(* IEC 61131-3 sources: JingjiangArm/moonboxpro_arm_8.4/Application/Application/任务列表/ExtTask/动作处理/油墨槽控制, 9 files *)

(* ---- StInkGrooveCtl.st ---- *)
(*@CES
Name=StInkGrooveCtl
Type=Gvl
TypeGuid=2db5746d-d284-4425-9f7f-2663a34b0ebc
Guid=c6ce6a04-2efb-4550-ab95-73592a3e1ea7
HasDeclaration=True
HasImplementation=False
*)
{DECLARATION}
TYPE StInkGrooveCtl :(*油墨槽控制@不保持|50bytes*)
STRUCT
	bySts							:BYTE;(*状态@就不用枚举了*)
	byMovingSts						:BYTE;(*运动状态|=0 不运动|=1 上升|=2 下降*)
	xCtlMode						:BOOL;(*控制模式|=false速度模式|=true 位置模式*)
	xMoveDir						:BOOL;(*运动的方向*)
	rVel							:REAL;(*速度值@r/min*)
	rMoveDis						:REAL;(*需要运动的距离@mm(带方向)*)
	diMoveDis_Pulse					:DINT;(*需要运动的距离(正值)@pulse*)
	wLastPulse_Act_Rd				:WORD;(*实际读取的脉冲数记录@上一拍*)
	xZeroValid						:BOOL;(*零位有效*)
	diPulse_Moved					:DINT;(*已经移动的脉冲|在原点处会更新为0*)
	rPos_Cur						:REAL;(*当前位置@mm|经过下限位零点后才有值*)
	iMsg							:TypeEnumInkGrooveMsg;(*信息 |=1 零点丢失
																  	 |=2 未确认基准
																   	 |=3 距离超限
																   	 |=4 上限位
																   	 |=5 下限位
																   	 |=6 速度模式下,运动异常*)
	diThisMovedPulse				:DINT;(*本次运动的距离@脉冲*)
	rThisMovedDis					:REAL;(*本次运动的距离@mm*)
	wLastPulse_Act_Rd_1				:WORD;(*实际读取的脉冲数记录@上一拍|用于计算本次运动的而距离值*)
	abyReseved						:ARRAY [1..11] OF BYTE;

END_STRUCT
END_TYPE

{IMPLEMENTATION}

(* ---- TypeEnumInkGrooveMsg.st ---- *)
(*@CES
Name=TypeEnumInkGrooveMsg
Type=Gvl
TypeGuid=2db5746d-d284-4425-9f7f-2663a34b0ebc
Guid=e4841006-6196-426e-9e86-ef53e879e515
HasDeclaration=True
HasImplementation=False
*)
{DECLARATION}
TYPE TypeEnumInkGrooveMsg :
(*信息枚举@和语言文件相关|1--9错误码|200以后为状态*)
(
	MSG_NONE:=0,(*无意义*)
	MSG_ZEROINVALID:=1,(*零点非法*)
	MSG_BASEINFINVALID,(*基准信息未确认*)
	MSG_MOVEDIS_OUTLIMTIT,(*运动距离超限*)
	MSG_UPLIMIT,(*上限位*)
	MSG_DNLIMIT,(*下限位*)
	MSG_MOVEFAILED,(*运动失败=6*)

	MSG_UPING:=200,(*向上运动中*)
	MSG_DNING(*向下运动中*)
);
END_TYPE

{IMPLEMENTATION}

(* ---- KS_BtnClick.st ---- *)
(*@CES
Name=KS_BtnClick
Type=FunctionBlock
TypeGuid=6f9dac99-8de1-4efc-8465-68ac443b7d08
Guid=4b1f190c-8fa5-4402-be53-ffd017a7b610
HasDeclaration=True
HasImplementation=True
*)
{DECLARATION}
FUNCTION KS_BtnClick : BOOL
(*按钮的单击双击长按处理*)
(*双击信号|在设定时间内按下2次输出信号*)
(*单击信号|第一次按下后超过i_iTime_ms时间未按下第二次按键输出单击事件,只有效一个周期*)
(*长按信号|第一次按下后超过i_iTime_ms时间未取消输出长按信号,直到松开*)
(*500ms还是有点感觉*)
VAR_INPUT
	i_xBtn:BOOL;
	i_wTime_ms:WORD:=300;(*时间*)
	i_byCycleTime_ms:BYTE:=20;(*周期时间*)
	i_pxClick:POINTER TO BOOL;(*单击有效(相当于按下等待i_wTime_ms时间后输出单击事件)@支持指针=0*)
	i_pxDoubleClick:POINTER TO BOOL;(*单击有效(相当于按下等待i_wTime_ms时间后输出单击事件)@支持指针=0*)
	i_pxHold:POINTER TO BOOL;(*按钮长按(相当于按下等待i_wTime_ms时间后输出单击事件)@支持指针=0*)
	i_pwCnt:POINTER TO WORD;(*时间周期计数|@./15作为按钮第一次按下沿标志
										  |@./14作为按钮第一次按下超时标志
										  |@./13作为按钮第一次按下抬起的标志
										  |@./12作为按钮第二次按下沿标志
										  |@故该值最大到16#FFF=4095*)
END_VAR
VAR
	wCnt: WORD;
	xDoubleClick:BOOL;
	xClick:BOOL;(*单击*)
	xHold:BOOL;(*长按*)
	xBtnU2D_1st: BOOL;(*按钮第一次按下沿标志*)
	xBtnU2DTimeOut_1st:BOOL;(*按钮第一次按下超时了*)
	xBtnD2U_1st: BOOL;(*按钮第一次按下到抬起标志*)
	xBtnU2D_2st: BOOL;(*按钮第二次抬起到按下沿标志*)
	wCnt_Use: WORD;(*实际计数值@最大16#fff*)
	xStopCnt: BOOL;(*停止计数标志*)
END_VAR
{IMPLEMENTATION}
IF i_pwCnt<>0 THEN
	wCnt:=i_pwCnt^;
END_IF
xBtnU2D_1st:=wCnt.15;
xBtnU2DTimeOut_1st:=wCnt.14;
xBtnD2U_1st:=wCnt.13;
xBtnU2D_2st:=wCnt.12;
wCnt_Use:=wCnt AND 16#FFF;(*只取低12bit*)

(*其实用状态机更好一些|有点乱*)
IF NOT xBtnU2D_1st THEN(*刚开始检测第一次按键*)
	IF i_xBtn THEN
		xBtnU2D_1st:=TRUE;
		(*标志初始化*)
		wCnt_Use:=0;
		xBtnU2DTimeOut_1st:=FALSE;
		xBtnD2U_1st:=FALSE;
		xBtnU2D_2st:=FALSE;
	END_IF
ELSE
	IF NOT xBtnD2U_1st THEN(*第一次的还没抬起来*)
		IF NOT i_xBtn THEN(*按钮抬起来了*)
			IF xBtnU2DTimeOut_1st THEN(*超过时间了@复位标志*)
				wCnt_Use:=0;
				xBtnU2DTimeOut_1st:=FALSE;
				xBtnU2D_1st:=FALSE;
				xStopCnt:=TRUE;(*停止计数*)
			ELSE(*未超过时间,继续检测*)
				xBtnD2U_1st:=TRUE;
			END_IF
		ELSE(*按下的时间太长了@输出长按标志*)
			(*超过时间了@复位标志*)
			IF NOT xBtnU2DTimeOut_1st THEN
				IF wCnt_Use*i_byCycleTime_ms>i_wTime_ms THEN
					wCnt_Use:=0;
					xBtnU2DTimeOut_1st:=TRUE;(*超时了*)
					xStopCnt:=TRUE;(*停止计数*)
					xHold:=TRUE;(*长按*)
				END_IF
			ELSE
				xStopCnt:=TRUE;(*停止计数*)
				xHold:=TRUE;(*长按*)
			END_IF
		END_IF
	ELSE
		IF NOT xBtnU2D_2st THEN(*第二次还未按下*)
			IF i_xBtn THEN(*再次按下*)
				IF wCnt_Use*i_byCycleTime_ms<=i_wTime_ms THEN(*在时间间隔内*)
					xDoubleClick:=TRUE;(*输出*)
				ELSE(*超过了时间|则不输出*)
					xDoubleClick:=FALSE;
				END_IF
				xBtnU2D_2st:=TRUE;(*第二次按下了*)
				xStopCnt:=TRUE;(*停止计数*)
			ELSE
				(*控制结束了*)
				IF wCnt_Use*i_byCycleTime_ms>i_wTime_ms THEN(*超过时间了@复位标志*)
					wCnt_Use:=0;
					xBtnU2D_1st:=FALSE;(*第一次按下复位*)
					xBtnD2U_1st:=FALSE;(*第一次抬起复位*)
					xStopCnt:=TRUE;(*停止计数*)
					xClick:=TRUE;(*输出单击事件*)
				END_IF
			END_IF
		ELSE(*第二次抬起按下了*)
			xStopCnt:=TRUE;(*停止计数*)
			IF NOT i_xBtn THEN(*抬起了,复位所有状态*)
				wCnt_Use:=0;
				xBtnU2D_1st:=FALSE;(*第一次按下复位*)
				xBtnD2U_1st:=FALSE;(*第一次抬起复位*)
				xBtnU2D_2st:=FALSE;(*第二次按下复位*)
			END_IF
		END_IF
	END_IF

	IF NOT xStopCnt THEN
		wCnt_Use:=wCnt_Use+1;(*计时开始*)
		IF wCnt_Use>=16#FFF THEN(*最大值限制*)
			wCnt_Use:=16#FFF;
		END_IF
	END_IF
END_IF

wCnt:=wCnt_Use;(*按位或*)
wCnt.15:=xBtnU2D_1st;
wCnt.14:=xBtnU2DTimeOut_1st;
wCnt.13:=xBtnD2U_1st;
wCnt.12:=xBtnU2D_2st;
IF i_pwCnt<>0 THEN
	i_pwCnt^:=wCnt;
END_IF
IF i_pxClick<>0 THEN
	i_pxClick^:=xClick;
END_IF
IF i_pxDoubleClick<>0 THEN
	i_pxDoubleClick^:=xDoubleClick;
END_IF
IF i_pxHold<>0 THEN
	i_pxHold^:=xHold;
END_IF

(* ---- KS_GetInkGrooveBaseInf.st ---- *)
(*@CES
Name=KS_GetInkGrooveBaseInf
Type=FunctionBlock
TypeGuid=6f9dac99-8de1-4efc-8465-68ac443b7d08
Guid=6496d967-7a0d-4af8-a414-ba22caa8f71e
HasDeclaration=True
HasImplementation=True
*)
{DECLARATION}
FUNCTION KS_GetInkGrooveBaseInf : BOOL
(*获取油墨槽基准信息*)
VAR_INPUT
	i_xEn:BOOL;(*获取使能@当前位置是有效的@且不在运动中*)
	i_xGetBtn:BOOL;(*获取按钮@沿触发*)
	i_rGirth:REAL;(*此时的版周长@mm*)
	i_rPos_Cur:REAL;(*此时位置@mm*)
	i_pxBaseInfValid:POINTER TO BOOL;(*基准信息有效*)
	i_prGirth_Base:POINTER TO REAL;(*基准周长(mm)@以该周长作为基准,计算其他周长的变化量*)
	i_prPos_Base:POINTER TO REAL;(*基准位置(mm)@基准周长对应的位置*)
END_VAR
VAR
END_VAR
{IMPLEMENTATION}
IF i_prGirth_Base<>0 AND
	i_prPos_Base<>0 THEN
	IF i_xEn THEN
		IF i_xGetBtn THEN
			i_pxBaseInfValid^:=TRUE;
			i_prGirth_Base^:=i_rGirth;
			i_prPos_Base^:=i_rPos_Cur;
		END_IF
	END_IF
END_IF

(* ---- KS_GetPulse_ActEx.st ---- *)
(*@CES
Name=KS_GetPulse_ActEx
Type=FunctionBlock
TypeGuid=6f9dac99-8de1-4efc-8465-68ac443b7d08
Guid=fa7aacb3-70fc-4571-89fd-f05cb3be533c
HasDeclaration=True
HasImplementation=True
*)
{DECLARATION}
FUNCTION KS_GetPulse_ActEx : INT(*读取实际的走了的脉冲数*)
(*2025.6.14.134137 增加累计取反*)
VAR_INPUT
	i_xRev:BOOL;(*取反标志|累计取反@2025.6.14.134133*)
	pwStepDrivePulse_Act_Rd :POINTER TO WORD;(*读取到的脉冲数*)
	pwStepDrivePulse_Act_Rd_Bak:POINTER TO WORD;(*上个周期读到的脉冲数*)
	pdiStepDrivePulse_Act:POINTER TO DINT;(*实际走的脉冲数*)
END_VAR
VAR
	iStepDrivePulse_Act_Rd: INT;
	iStepDrivePulse_Act_Rd_Bak: INT;
	iDeltaPulse: INT;(*步进电机脉冲变化量*)
END_VAR
{IMPLEMENTATION}
KS_GetPulse_ActEx:=0;
IF pwStepDrivePulse_Act_Rd<>0 AND pwStepDrivePulse_Act_Rd_Bak<>0 AND pdiStepDrivePulse_Act <>0 THEN;
ELSE
	KS_GetPulse_ActEx:=-1;
	RETURN;
END_IF

iStepDrivePulse_Act_Rd:=WORD_TO_INT(pwStepDrivePulse_Act_Rd^);
iStepDrivePulse_Act_Rd_Bak:= WORD_TO_INT(pwStepDrivePulse_Act_Rd_Bak^);

IF iStepDrivePulse_Act_Rd <> iStepDrivePulse_Act_Rd_Bak THEN
	iDeltaPulse:=(iStepDrivePulse_Act_Rd-iStepDrivePulse_Act_Rd_Bak);
	IF i_xRev THEN
		iDeltaPulse:=-iDeltaPulse;
	END_IF
	pdiStepDrivePulse_Act^:=pdiStepDrivePulse_Act^+iDeltaPulse;
ELSE;
END_IF

pwStepDrivePulse_Act_Rd_Bak^:=INT_TO_WORD(iStepDrivePulse_Act_Rd);(*保存上个周期的值*)

(* ---- KS_InkGrooveCtl_1Axis.st ---- *)
(*@CES
Name=KS_InkGrooveCtl_1Axis
Type=FunctionBlock
TypeGuid=6f9dac99-8de1-4efc-8465-68ac443b7d08
Guid=2dac3483-8274-459a-981e-f455ba92ec89
HasDeclaration=True
HasImplementation=True
*)
{DECLARATION}
FUNCTION KS_InkGrooveCtl_1Axis : BOOL
(*油墨槽控制函数@单轴*)
(*根据按钮控制输出*)
(*走定位是按照速度模式+位置模式输出处理@因为位置模式目前架构只支持最多65535脉冲*)
(*我们定义正值是向上运动的|默认方式是向上运动的,可以通过i_xMoveDirRev输入切换方向*)
VAR_INPUT
	i_xEn:BOOL;(*控制使能*)
	i_xCanMove:BOOL;(*可以运动标志@例如非急停*)
	i_xClrMsg:BOOL;(*清除msg*)
	i_lrDis_1Pulse:REAL;(*单位脉冲对应的距离@mm/pulse*)
	i_iCycleTime_Plc:INT:=20;(*程序周期时间@ms*)
	i_rGirth:REAL;(*当前版周长@mm*)
	i_xBaseInfValid:BOOL;(*基准信息是有效的*)
	i_rGirth_Base:REAL;(*基准周长(mm)@以该周长作为基准,计算其他周长的变化量*)
	i_rPos_Base:REAL;(*基准位置(mm)@基准周长对应的位置*)
	i_xMoveDirRev:BOOL;(*运动方向取反*)
	i_xUp:BOOL;(*上升@长有效*)
	i_xUplimt:BOOL;(*上限位@硬件*)
	i_xDn:BOOL;(*下降@长有效*)
	i_xDn_Auto:BOOL;(*自动下降@沿触发(下降到i_xZeroSig位置)*)
	i_xDnlimt:BOOL;(*下限位@硬件|作为0点*)
	i_xUpClick : BOOL ;(*上升单击停止事件*)
	i_xDnClick : BOOL ;(*下降单击停止事件*)
	i_xToTarPos_Auto:BOOL;(*一键到位@沿触发*)
	i_xZeroSig:BOOL;(*零点信号(外部沿触发)@目前配置为下限位*)
	i_rSetVel:REAL;(*设置的运动速度@r/min*)
(*	i_diThisMovePulse:DINT;(*本次运动的脉冲@外部输入,就不在里面运算了*)*)
	i_rMaxMoveDis:REAL;(*最大运动距离@mm*)
	(*反馈*)
	i_wPulse_Act_Rd:WORD;(*读取的脉冲输出个数@用于计算当前位置*)
	i_xInPos:BOOL;(*到位标志@位置模式下反馈的标志*)
	i_xMoving_Act:BOOL;(*实际处于运动状态@再运动的时候就不能响应io*)
	i_xVelMode_MoveFailed:BOOL;(*速度模式下|运动失败了*)
	i_pstStInkGrooveCtl:POINTER TO StInkGrooveCtl;
(*
	(*输出@提供给脉冲输出函数处理*)
	i_pbySts:POINTER TO BYTE;(*状态@就不用枚举了|0 空闲
												|1 监控按钮*)
	i_pbyMovingSts:POINTER TO BYTE;(*运动状态|=0 不运动|=1 上升|=2 下降*)
	i_pxCtlMode:POINTER TO BOOL;(*控制模式|=false速度模式|=true 位置模式*)
	i_pxMoveDir:POINTER TO BOOL;(*运动的方向*)
	i_prVel:POINTER TO REAL;(*速度值@r/min*)
	i_prMoveDis:POINTER TO REAL;(*需要运动的距离@mm*)
	i_pwLastPulse_Act_Rd:POINTER TO WORD;(*实际读取的脉冲数记录@上一拍*)
	i_pxZeroValid:POINTER TO BOOL;(*零位有效*)
	i_pdiPulse_Moved:POINTER TO DINT;(*已经移动的脉冲|在原点处会更新为0*)
	i_prPos_Cur:POINTER TO REAL;(*当前位置@mm|经过下限位零点后才有值*)
	i_pbyMsg:POINTER TO BYTE;(*信息|=1 零点丢失
								   |=2 未确认基准
								   |=3 距离超限*)
*)
END_VAR
VAR
	lrPulse2Dis: LREAL;(*脉冲转换为距离系数@mm/pul*)
	bySts: BYTE;(*状态@就不用枚举了*)
	byMovingSts:BYTE;(*运动状态|=0 不运动|=1 上升|=2 下降*)
	xCtlMode:BOOL;(*控制模式|=FALSE速度模式|=TRUE 位置模式*)
	xMoveDir:BOOL;(*运动的方向*)
	rVel:REAL;(*速度值@r/min*)
	wPulseNum:WORD;(*位置模式脉冲个数@目前的逻辑只支持word输出*)
	rMoveDis:REAL;(*需要运动的距离@mm*)
	diMoveDis_Pulse: DINT;(*需要运动的距离@PULSE*)
	wLastPulse_Act_Rd:WORD;(*实际读取的脉冲数记录@上一拍*)
	diPulse_Moved:DINT;(*本次运动已经移动的脉冲|重新启动运动会更新*)
	rPos_Cur:REAL;(*当前位置@mm|经过下限位零点*)
	xZeroValid: BOOL;(*零位有效*)
	rSetVel:REAL;(*设置的运动速度@r/min*)
	rSetPos: REAL;(*设置的位置值mm*)
	xUpLimt_Use: BOOL;(*应用的上限位标志*)
	xDnLimt_Use: BOOL;(*应用的下限位标志*)
	diPluse_Act: DINT;(*相对零位走的脉冲数*)
(*	byMsg: BYTE;(*信息*)*)
	iMsg: TypeEnumInkGrooveMsg;(*信息*)
	diThisMovedPulse: DINT;(*本次运动的距离@脉冲*)
	wLastPulse_Act_Rd_1: WORD;(*用于计算本次运动距离*)
	rThisMovedDis: REAL;(*本次运动的距离@mm*)
	rPI:REAL:=3.1415926;
END_VAR
{IMPLEMENTATION}
IF i_pstStInkGrooveCtl<>0 THEN;
ELSE
	RETURN;
END_IF
IF i_xEn THEN

	bySts:=i_pstStInkGrooveCtl^.bySts;
	byMovingSts:=i_pstStInkGrooveCtl^.byMovingSts;
	rMoveDis:=i_pstStInkGrooveCtl^.rMoveDis;
	wLastPulse_Act_Rd:=i_pstStInkGrooveCtl^.wLastPulse_Act_Rd;
	diPulse_Moved:=i_pstStInkGrooveCtl^.diPulse_Moved;
	rPos_Cur:=i_pstStInkGrooveCtl^.rPos_Cur;
	xZeroValid:=i_pstStInkGrooveCtl^.xZeroValid;
	iMsg:=i_pstStInkGrooveCtl^.iMsg;

	diThisMovedPulse:=i_pstStInkGrooveCtl^.diThisMovedPulse;
	wLastPulse_Act_Rd_1:=i_pstStInkGrooveCtl^.wLastPulse_Act_Rd_1;

	(*脉冲转换为距离@mm*)
	IF i_lrDis_1Pulse<>0 THEN
		lrPulse2Dis:=i_lrDis_1Pulse;(*单个脉冲的距离@mm/pul*)
	ELSE
		lrPulse2Dis:=0.0002;
	END_IF

	(*计算本次走的脉冲数*)
	KS_GetPulse_ActEx(i_xMoveDirRev,
					ADR(i_wPulse_Act_Rd),
				 	ADR(wLastPulse_Act_Rd_1),
					ADR(diThisMovedPulse));
(*	diThisMovedPulse:=i_diThisMovePulse;*)
	rThisMovedDis:=diThisMovedPulse*lrPulse2Dis;

	(*距离计算*)
	(*计算实际走的脉冲数*)
	(*输出方向取反的时候 累计函数也要取反@2025.6.14.134430+*)
	KS_GetPulse_ActEx(i_xMoveDirRev,
					ADR(i_wPulse_Act_Rd),
				 	ADR(wLastPulse_Act_Rd),
					ADR(diPulse_Moved));

	(*零点信号检查*)
	IF i_xZeroSig THEN(*0点信号触发了*)
		xZeroValid:=TRUE;(*触发以后就不清除*)
		diPulse_Moved:=0;
		wLastPulse_Act_Rd:=i_wPulse_Act_Rd;
	END_IF

	IF xZeroValid THEN(*零位有效了@根据当前统计的脉冲数计算*)
		rPos_Cur:=diPulse_Moved*lrPulse2Dis;(*当前位置@mm*)
	ELSE(*没有零位的时候当前位置=0*)
		rPos_Cur:=0;
	END_IF

	(*动作实现*)
	rSetVel:=i_rSetVel;
	xUpLimt_Use:=i_xUplimt;
	xDnLimt_Use:=i_xDnlimt;

	IF NOT i_xCanMove THEN
		bySts:=0;(*空闲态*)
	ELSE(*可以运动的时候监控按钮*)
		IF bySts=0 THEN(*空闲时候检查*)
			IF i_xMoving_Act THEN(*处于运动中|不允许处理io信号*)
				i_xUp:=FALSE;
				i_xDn:=FALSE;
				i_xToTarPos_Auto:=FALSE;
				i_xDn_Auto:=FALSE;
			END_IF

			IF i_xUp THEN(*上升*)
				iMsg:=MSG_NONE;
				IF NOT xUpLimt_Use THEN(*未到限位*)
					bySts:=1;
				ELSE
					iMsg:=MSG_UPLIMIT;
				END_IF
			ELSIF i_xDn THEN(*下降*)
				iMsg:=MSG_NONE;
				IF NOT xDnLimt_Use THEN(*未到限位*)
					bySts:=2;
				ELSE
					iMsg:=MSG_DNLIMIT;
				END_IF
			ELSIF i_xToTarPos_Auto THEN(*一键自动到位*)
				iMsg:=MSG_NONE;
				IF xZeroValid THEN(*有0位才可以执行*)
					IF i_xBaseInfValid THEN
						rSetPos:=i_rGirth/2/rPI-i_rGirth_Base/2/rPI;(*和基准变化的位置-半径差@mm*)
						rSetPos:=-rSetPos;(*正值,需要油墨槽向下运动@处理方向*)
						rSetPos:=i_rPos_Base+rSetPos-rPos_Cur;(*计算相对当前位置的增量*)
						IF rSetPos>0 THEN(*正值@向上运动*)
							IF NOT xUpLimt_Use THEN(*未到限位*)
								bySts:=10;
							ELSE
								iMsg:=MSG_UPLIMIT;
							END_IF
						ELSIF rSetPos<0 THEN(*负值@向下运动*)
							IF NOT xDnLimt_Use THEN(*未到限位*)
								bySts:=10;
							ELSE
								iMsg:=MSG_DNLIMIT;
							END_IF
						END_IF
					ELSE(*未确认基准*)
						iMsg:=MSG_BASEINFINVALID;
					END_IF
				ELSE(*没有零位*)
					iMsg:=MSG_ZEROINVALID;
				END_IF
			ELSIF i_xDn_Auto THEN(*自动下降*)
				iMsg:=MSG_NONE;
				diThisMovedPulse:=0;(*本次运动的距离清零*)
				IF NOT xDnLimt_Use THEN(*未到限位*)
					bySts:=20;
				ELSE
					iMsg:=MSG_DNLIMIT;
				END_IF
			END_IF
		END_IF
	END_IF
	(*信息清理*)
	IF iMsg<>MSG_NONE THEN
		IF i_xClrMsg THEN
			iMsg:=MSG_NONE;
		END_IF
	END_IF

	rVel:=rSetVel;(*设置的速度值*)
	CASE bySts OF
		0:;(*空闲时候@啥都不干*)
			byMovingSts:=0;
			rMoveDis:=0;
		1,2:(*手动上升\下降*)
			xCtlMode:=FALSE;(*速度模式*)
			rMoveDis:=0;(*设置的位置值*)
			IF bySts=1 THEN
				IF NOT i_xUp THEN(*取消上升*)
					bySts:=0;
				END_IF
				byMovingSts:=1;(*上升*)
			ELSE
				IF NOT i_xDn THEN(*取消上升*)
					bySts:=0;
				END_IF
				byMovingSts:=2;(*下降*)
			END_IF

			diThisMovedPulse:=0;(*本次运动的距离清零*)
		10:(*一键到位@速度模式+位置模式|将速度参数和位置参数都下发下去*)
			xCtlMode:=TRUE;(*按照位置模式输出*)
			rMoveDis:=rSetPos;(*设置的位置值*)
			IF rMoveDis>0 THEN
				byMovingSts:=1;(*上升*)
			ELSE
				byMovingSts:=2;(*下降*)
			END_IF
			bySts:=11;
			diThisMovedPulse:=0;(*本次运动的距离清零*)
		11:(*等待运动完成*)
			xCtlMode:=TRUE;(*按照位置模式输出*)
			(*rMoveDis@保持case10中的值*)
			IF i_xInPos OR (*到位标志|退出case*)
				i_xUp OR i_xDn  OR i_xUpClick  THEN(*上升或者下降按钮被按下则取消运动*)
				bySts:=0;
			END_IF
			(*运动的距离超限了,就停止吧*)
			IF ABS(rThisMovedDis)>ABS(i_rMaxMoveDis) THEN
				bySts:=0;
			END_IF

		20:(*自动下降到下限位@按照速度模式一直向下运动直到触发限位或者运动了最大距离*)
			xCtlMode:=FALSE;(*按照速度模式输出*)
			rMoveDis:=0;(*设置的位置值*)
			byMovingSts:=2;(*下降*)
			IF xDnLimt_Use OR(*到达下限位了*)
				i_xUp OR i_xDn OR i_xDnClick THEN(*上升或者下降按钮被按下则取消运动*)
				bySts:=0;
			END_IF
			(*运动的距离超限了,就停止吧*)
			IF ABS(rThisMovedDis)>ABS(i_rMaxMoveDis) THEN
				bySts:=0;
			END_IF
	ELSE
		bySts:=0;
		byMovingSts:=0;
		rMoveDis:=0;
	END_CASE
	IF bySts = 0 THEN(*退出状态时候|复位运动状态@使用case清除会滞后一个周期*)
		byMovingSts:= 0;
	END_IF

	diMoveDis_Pulse:=LREAL_TO_DINT(rMoveDis/lrPulse2Dis);(*将位置转换为脉冲*)
	(*方向处理*)
	IF byMovingSts=1 THEN(*上升*)
		xMoveDir:=FALSE;
	ELSIF byMovingSts =2 THEN(*下降*)
		xMoveDir:=TRUE;
	ELSE;(*保持之前的*)
	END_IF
	(*方向取反控制*)
	IF i_xMoveDirRev THEN
		xMoveDir:=NOT xMoveDir;
	END_IF

	(*使能时限位处理@一直检查*)
	IF byMovingSts<>0 THEN
		IF byMovingSts=1 THEN(*上升检查一下上限位*)
			IF xUpLimt_Use THEN
				iMsg:=MSG_UPLIMIT;(*到限位信息提示*)
				byMovingSts:=0;
			ELSE
				iMsg:=MSG_UPING;(*输出上升中*)
			END_IF
		END_IF
		IF byMovingSts=2 THEN(*下降检查一下下限位*)
			IF xDnLimt_Use THEN
				iMsg:=MSG_DNLIMIT;(*到限位信息提示*)
				byMovingSts:=0;
			ELSE
				iMsg:=MSG_DNING;(*输出下降中*)
			END_IF
		END_IF

		(*2025.6.10.151223+*)
		IF i_xVelMode_MoveFailed THEN
			iMsg:=MSG_MOVEFAILED;
		END_IF
	ELSE;(*功能的特性,会将设置值全部清0*)
		(*如果处于运动中退出,就将信息清除*)
		IF iMsg=MSG_UPING OR iMsg=MSG_DNING THEN
			iMsg:=MSG_NONE;
		END_IF
	END_IF
ELSE
	wLastPulse_Act_Rd:=i_wPulse_Act_Rd;
	wLastPulse_Act_Rd_1:=i_wPulse_Act_Rd;
END_IF

(*指针处理*)
i_pstStInkGrooveCtl^.bySts:=bySts;
i_pstStInkGrooveCtl^.byMovingSts:=byMovingSts;
i_pstStInkGrooveCtl^.xCtlMode:=xCtlMode;
i_pstStInkGrooveCtl^.xMoveDir:=xMoveDir;
i_pstStInkGrooveCtl^.rVel:=rVel;
i_pstStInkGrooveCtl^.rMoveDis:=rMoveDis;
i_pstStInkGrooveCtl^.diMoveDis_Pulse:=ABS(diMoveDis_Pulse);(*只保留正值@方向由标志控制*)
i_pstStInkGrooveCtl^.wLastPulse_Act_Rd:=wLastPulse_Act_Rd;
i_pstStInkGrooveCtl^.diPulse_Moved:=diPulse_Moved;
i_pstStInkGrooveCtl^.rPos_Cur:=rPos_Cur;
i_pstStInkGrooveCtl^.xZeroValid:=xZeroValid;
i_pstStInkGrooveCtl^.iMsg:=iMsg;
i_pstStInkGrooveCtl^.diThisMovedPulse:=diThisMovedPulse;
i_pstStInkGrooveCtl^.wLastPulse_Act_Rd_1:=wLastPulse_Act_Rd_1;
i_pstStInkGrooveCtl^.rThisMovedDis:=rThisMovedDis;

(* ---- KS_PulseOutCtl.st ---- *)
(*@CES
Name=KS_PulseOutCtl
Type=FunctionBlock
TypeGuid=6f9dac99-8de1-4efc-8465-68ac443b7d08
Guid=26372ce9-281b-45a3-9b8d-535af9137d46
HasDeclaration=True
HasImplementation=True
*)
{DECLARATION}
FUNCTION KS_PulseOutCtl : INT
(*2025.2.19.105619 脉冲输出控制函数@主要针对1610模块以及新款16d驱动器io*)
(*切换模式的话,需要取消使能|i_pbyOutSts^=3只有速度模式才会被写入*)
VAR_INPUT
	i_xEn:BOOL;(*控制使能了*)
	i_xClrPulse_Act_Rd:BOOL;(*清理实际的脉冲数*)
	i_byJudgeOutsts_WaitNum:BYTE:=10;(*等待周期数@超过该值强制清除输出中标志|时间=i_byJudgeOutsts_WaitNum*执行周期*)
	i_dwPulse_1r:DWORD;(*一圈的脉冲数*)
	i_xCtlMode:BOOL;(*控制模式@=false 速度模式|=true 位置模式*)
	i_xVelMod_Run:BOOL;(*速度模式下,启动运动标志@前提是状态机已经启动到了脉冲输出case*)
	i_xDir:BOOL;(*输出的方向@false=正向|=true 反向*)
	i_rVel_Sa:REAL;(*起始速度@r/min*)
	i_rVel:REAL;(*速度值@速度模式 r/min*)
	i_iAccTime_ms:INT;(*加速时间@100*)(*ms*)
	i_pwPulse:POINTER TO WORD;(*输出的脉冲个数-写入后就清零了@位置模式*)
	(*反馈信号*)
	i_xPulseOutting_Rd:BOOL;(*读取到的脉冲输出中标志*)
	i_wPulse_Act_Rd:WORD;(*读取的脉冲输出个数*)
	(*输出*)
	i_piState			:POINTER TO TypeEnumStepDriveStat;(*控制状态@状态机标志*)
	i_pwCtlBit_Wr		:POINTER TO WORD;(*控制bit写入*)
	i_pwFre_Sa_Wr		:POINTER TO WORD;(*起始频率写入到模块或者驱动器的值*)
	i_pwFreq_Tar_Wr		:POINTER TO WORD;(*目标频率写入到模块或者驱动器的值*)
	i_pwAccSaToTar_Wr	:POINTER TO WORD;(*频率加速度写入到模块或者驱动器的值*)
	i_pwPulse_Pos_Wr	:POINTER TO WORD;(*脉冲数写入到模块或者驱动器的值*)
	i_pdiPluse_Act		:POINTER TO DINT;(*实际的脉冲数@开始的时候会清除*)
	i_pwLastPulse_Act_Rd:POINTER TO WORD;(*实际读取的脉冲数记录@上一拍*)
	i_pbyOutSts			:POINTER TO BYTE;(*输出状态|=0 不输出|=1 输出@逻辑|=2反馈正在运行|=3异常|=255 准备写入@进入case*)
	i_pxCtlMod_Cur		:POINTER TO BOOL;(*当前控制模式@=false 速度模式|=true 位置模式*)
	i_pbyWaitCnt		:POINTER TO BYTE;(*周期等待计数@根据程序周期计算等待时间*)
END_VAR
VAR
	lrTemp:LREAL;
	dwPulse_Pos:DWORD;(*目前只取了word@因为模块和驱动器都只支持到word类型*)
	lrFreq_Sa: LREAL;(*起始频率@P/S*)
	lrFreq_Tar: LREAL;(*目标频率@P/S*)
	lrAccSaToTar:LREAL;(*起始频率加速到目标频率的加速度@hz/s*)
	wFre_Sa_Wr: WORD;(*起始频率写入到模块或者驱动器的值*)
	wFreq_Tar_Wr: WORD;(*目标频率写入到模块或者驱动器的值*)
	wAccSaToTar_Wr: WORD;(*频率加速度写入到模块或者驱动器的值*)
	wPulse_Pos_Wr:WORD;(*脉冲数写入到模块或者驱动器的值*)
	iState: TypeEnumStepDriveStat;(*控制状态机*)
	wCTLBit: WORD;(*控制位*)
	diPluse_Act:DINT;(*实际的脉冲数*)
	wLastPulse_Act_Rd:WORD;(*实际读取的脉冲数记录@上一拍*)
	iAccTime_ms: INT;
	byOutSts: BYTE;(*输出状态|=0 不输出|=1 输出|=2异常*)
	xCtlMod_Cur: BOOL;(*当前控制模式@=false 速度模式|=true 位置模式*)
	byWaitCnt: BYTE;(*周期等待计数*)

	xFreq_Sa_Wr:BOOL;(*启动频率写入标志*)
	xFreq_Tar_Wr:BOOL;(*目标频率写入标志*)
	xFreq_AccSaToTar_Wr:BOOL;(*加速度频率写入标志*)
	xFreq_Pulse_Pos_Wr:BOOL;(*脉冲写入标志*)
END_VAR
VAR CONSTANT
(*
bit9:反馈脉冲数清零
bit10:脉冲输出标志，1：输出中
bit11:电机方向
bit12:速度模式时，高电平输出脉冲，低电平停止输出
bit13:位置模式时，上升沿开始输出脉冲，脉冲个数到达时停止输出
bit14:速度、位置模式 0：速度模式，1：位置模式
bit15:模块使能 0：脉冲输出无效，1：有效
*)
	c_wPosbak_Clear		:WORD:=16#0200;(*反馈脉冲数清零*)
	c_wStepDrive_Dir		:WORD:=16#0800;(*电机方向*)
	c_wSpeedMode_OutCtl	:WORD:=16#1000;(*速度模式输出控制*)
	c_wPosMode_OutCtl	:WORD:=16#2000;(*位置模式输出控制*)
	c_wPosMode			:WORD:=16#4000;(*默认为速度模式，有效为位置模式; 位置模式 速度模式选择，*)
	c_wAIModule_Valid		:WORD:=16#8000;(*模块使能*)
END_VAR
{IMPLEMENTATION}
IF i_pdiPluse_Act<>0 THEN
	diPluse_Act:=i_pdiPluse_Act^;
END_IF
IF i_pwLastPulse_Act_Rd<>0 THEN
	wLastPulse_Act_Rd:=i_pwLastPulse_Act_Rd^;
END_IF

IF i_xEn THEN
	(*写入到模块或者驱动器的值*)
	IF i_pwPulse<>0 THEN(*写入的脉冲数*)
		wPulse_Pos_Wr:=i_pwPulse^;
	END_IF
	IF i_piState<>0 THEN
		iState:=i_piState^;
	END_IF
	IF i_pbyOutSts<>0 THEN
		byOutSts:=i_pbyOutSts^;
	END_IF
	IF i_pxCtlMod_Cur<>0 THEN
		xCtlMod_Cur:=i_pxCtlMod_Cur^;
	END_IF
	IF i_pbyWaitCnt<>0 THEN
		byWaitCnt:=i_pbyWaitCnt^;
	END_IF

	IF i_iAccTime_ms<>0 THEN
		iAccTime_ms:=ABS(i_iAccTime_ms);
	ELSE
		iAccTime_ms:=100;
	END_IF
	lrTemp:=EXPT(2,12)/EXPT(5,6);(*由EXPT(2,18)/EXPT(10,6)化简而来*)
	(*将起始速度转换为频率*)
	lrFreq_Sa:=i_dwPulse_1r*ABS(i_rVel_Sa)/60.0;(*pul/s*)
	(*将目标速度转换为频率*)
	lrFreq_Tar:=i_dwPulse_1r*ABS(i_rVel)/60.0;(*pul/s*)

	(*起始频率大于目标频率时 让起始频率等于目标频率*)
	IF lrFreq_Sa>lrFreq_Tar THEN
		lrFreq_Sa:=lrFreq_Tar;
	END_IF
	(*计算起始频率应该写入的值*)
	wFre_Sa_Wr:=LREAL_TO_WORD(lrFreq_Sa*lrTemp);(*计算写入模块中的值*)

	(*计算目标频率应该写入的值*)
	wFreq_Tar_Wr:=LREAL_TO_WORD(lrFreq_Tar*lrTemp);(*计算写入模块中的值*)

(*计算加速度*)
	lrTemp:=EXPT(2,22)/EXPT(5,12);(*EXPT(2,32)/EXPT(10,12)化简得到的*)(*计算出的加速度*该值就是需要写入模块中的值*)
	(*计算加速度@从起始频率到目标频率的加速度*)
	lrAccSaToTar:=ABS(lrFreq_Tar-lrFreq_Sa)*1000/iAccTime_ms;(*HZ/S*)
	(*需要写入到模块中的加速度值*)
	wAccSaToTar_Wr:=LREAL_TO_WORD(lrAccSaToTar*lrTemp);

	(*启动case*)
	IF iState = STEPDRIVE_IDLE THEN
		iState:=STEPDRIVE_RUN;
	END_IF
	wCTLBit:=0;(*清零该控制位*)
	xFreq_Sa_Wr:=FALSE;
	xFreq_Tar_Wr:=FALSE;
	xFreq_AccSaToTar_Wr:=FALSE;
	xFreq_Pulse_Pos_Wr:=FALSE;
	CASE iState OF
	STEPDRIVE_IDLE:;
	STEPDRIVE_RUN,STEPDRIVE_CLR:
		IF i_xClrPulse_Act_Rd THEN
			wCTLBit:=c_wPosbak_Clear;
		END_IF
		iState:=STEPDRIVE_WAITING;
		(*放在这个周期是希望在计数清零执行后*)
		diPluse_Act:=0;(*初始化脉冲计数值*)
		wLastPulse_Act_Rd:=i_wPulse_Act_Rd;(*初始化上个周期的值*)
		byOutSts:=255;
		xCtlMod_Cur:=i_xCtlMode;
		byWaitCnt:=0;
	STEPDRIVE_WAITING:(*等一个周期*)
		iState:=STEPDRIVE_MODULE_VALID;
	STEPDRIVE_MODULE_VALID:(*模块使能*)
		(*放在这个周期是希望在计数清零执行后*)
		diPluse_Act:=0;(*初始化脉冲计数值*)
		wLastPulse_Act_Rd:=i_wPulse_Act_Rd;(*初始化上个周期的值*)

		wCTLBit:=c_wAIModule_Valid;
		IF xCtlMod_Cur THEN (*位置模式*)
			wCTLBit:=wCTLBit+c_wPosMode;
		ELSE(*速度模式*)
			wCTLBit:=wCTLBit;
		END_IF

		IF i_xDir THEN (*步进电机方向*)
			wCTLBit:=wCTLBit+c_wStepDrive_Dir;
		ELSE;(*默认方向*)
		END_IF
		(*2022.11.19.160459 从case-STEPDRIVE_PULSEOUT复制到此处 提前写入一个周期
		@发现手动有时候脉冲输出不对
		@发现手动有时候会步输出。测试复制到此处出现的概率小很多了*)
		(*写入启动频率 目标频率 加速度值*)
		xFreq_Sa_Wr:=TRUE;(*启动频率写入标志*)
		xFreq_Tar_Wr:=TRUE;(*目标频率写入标志*)
		xFreq_AccSaToTar_Wr:=TRUE;(*加速度值写入标志*)
		iState:=STEPDRIVE_PULSEOUT;(*进入脉冲输出逻辑*)
	STEPDRIVE_PULSEOUT:(*脉冲输出*)(*脉冲输出比电机方向配置晚一个周期*)
		(*写入启动频率 目标频率 加速度值*)
		xFreq_Sa_Wr:=TRUE;(*启动频率写入标志*)
		xFreq_Tar_Wr:=TRUE;(*目标频率写入标志*)
		xFreq_AccSaToTar_Wr:=TRUE;(*加速度值写入标志*)

		IF xCtlMod_Cur THEN (*位置模式*)
			wCTLBit:=c_wAIModule_Valid+c_wPosMode;
			(*写入脉冲数*)
			IF byOutSts=255 THEN(*未输出的时候才能写入*)
				IF wPulse_Pos_Wr<>0 THEN
					xFreq_Pulse_Pos_Wr:=TRUE;(*脉冲数写入标志*)
					wCTLBit:=wCTLBit+c_wPosMode_OutCtl;(*有效之后输出脉冲*)(*上升沿触发*)
					byOutSts:=1;(*置位输出中标志*)
					byWaitCnt:=0;
				END_IF
			ELSIF byOutSts=1 THEN(*输出中*)
				IF byWaitCnt>=i_byJudgeOutsts_WaitNum THEN(*超过计时@判断是否结束|认为超过这个时间肯定运动了*)
					IF NOT i_xPulseOutting_Rd THEN
						byOutSts:=255;
					END_IF
				ELSE(*等待*)
					byWaitCnt:=byWaitCnt+1;
					IF i_xPulseOutting_Rd THEN
						byOutSts:=2;
					END_IF
				END_IF
			ELSIF byOutSts=2 THEN(*实际也运行了*)
				IF NOT i_xPulseOutting_Rd THEN
					byOutSts:=255;
				END_IF
			END_IF
		ELSE(*速度模式*)(*该模式启动之后就不能更改参数，除非重新开始*)
			wCTLBit:=c_wAIModule_Valid;
			IF byOutSts=255 THEN(*未输出的时候才能写入*)
				IF i_xVelMod_Run THEN
					wCTLBit:=wCTLBit+c_wSpeedMode_OutCtl;(*有效之后输出脉冲*)
					byOutSts:=1;(*置位输出中标志*)
					byWaitCnt:=0;
				END_IF
			ELSE
				wCTLBit:=wCTLBit+c_wSpeedMode_OutCtl;
				IF byOutSts=1 THEN(*输出中*)
					IF byWaitCnt>=i_byJudgeOutsts_WaitNum THEN(*超过计时@判断是否结束|认为超过这个时间肯定运动了*)
						IF NOT i_xPulseOutting_Rd THEN
							IF NOT i_xVelMod_Run THEN(*退出运动了*)
								byOutSts:=255;
							ELSE(*还未执行运动则报错*)
								byOutSts:=3;
							END_IF
						ELSE(*实际运动了*)
							byOutSts:=2;
						END_IF
					ELSE(*等待*)
						byWaitCnt:=byWaitCnt+1;
						IF i_xPulseOutting_Rd THEN(*已经再运行了*)
							byOutSts:=2;
						END_IF
					END_IF
				ELSIF byOutSts=2 THEN(*实际确实再运行了*)
					IF NOT i_xVelMod_Run AND NOT i_xPulseOutting_Rd THEN(*退出运动了*)
						byOutSts:=255;
					END_IF
				ELSE(*byOutSts=3*)
					IF NOT i_xVelMod_Run THEN(*退出运动了*)
						byOutSts:=255;
					END_IF
				END_IF
			END_IF
		END_IF

		IF i_xDir THEN (*步进电机方向*)
			wCTLBit:=wCTLBit+c_wStepDrive_Dir;
		ELSE;(*默认方向*)
		END_IF
	STEPDRIVE_ALARM:;(*报警步*)
	ELSE;
	END_CASE

	(*计算本次实际走的脉冲数*)
	KS_GetPulse_Act(ADR(i_wPulse_Act_Rd),
				 	ADR(wLastPulse_Act_Rd),
					ADR(diPluse_Act));
ELSE(*不使能*)
	iState:=STEPDRIVE_IDLE;
	wPulse_Pos_Wr:=0;(*写入的脉冲为0*)
	IF i_xPulseOutting_Rd THEN
		byOutSts:=1;
	ELSE
		byOutSts:=0;
	END_IF
END_IF

(*输出*)
IF i_pwCtlBit_Wr<>0 THEN
	i_pwCtlBit_Wr^:=wCTLBit;
END_IF
IF i_piState<>0 THEN
	i_piState^:=iState;
END_IF
IF i_pwFre_Sa_Wr<>0 THEN
	IF xFreq_Sa_Wr THEN(*启动频率写入*)
		i_pwFre_Sa_Wr^:=wFre_Sa_Wr;
	ELSE
		i_pwFre_Sa_Wr^:=0;
	END_IF
END_IF
IF i_pwFreq_Tar_Wr<>0 THEN
	IF xFreq_Tar_Wr THEN(*目标频率写入*)
		i_pwFreq_Tar_Wr^:=wFreq_Tar_Wr;
	ELSE
		i_pwFreq_Tar_Wr^:=0;
	END_IF
END_IF
IF i_pwAccSaToTar_Wr<>0 THEN
	IF xFreq_AccSaToTar_Wr THEN(*加速度写入*)
		i_pwAccSaToTar_Wr^:=wAccSaToTar_Wr;
	ELSE
		i_pwAccSaToTar_Wr^:=0;
	END_IF
END_IF
IF i_pwPulse_Pos_Wr<>0 THEN
	IF xFreq_Pulse_Pos_Wr THEN(*脉冲写入*)
		i_pwPulse_Pos_Wr^:=wPulse_Pos_Wr;
		wPulse_Pos_Wr:=0;(*脉冲写入后就写0*)
	ELSE
		i_pwPulse_Pos_Wr^:=0;
	END_IF
END_IF

IF i_pdiPluse_Act<>0 THEN
	i_pdiPluse_Act^:=diPluse_Act;
END_IF
IF i_pwLastPulse_Act_Rd<>0 THEN
	i_pwLastPulse_Act_Rd^:=wLastPulse_Act_Rd;
END_IF
(*注意顺序i_pwPulse_Pos_Wr 写入之后*)
IF i_pwPulse<>0 THEN(*写入的脉冲数*)
	i_pwPulse^:=wPulse_Pos_Wr;
END_IF

IF i_pbyOutSts<>0 THEN
	i_pbyOutSts^:=byOutSts;
END_IF
IF i_pxCtlMod_Cur<>0 THEN
	i_pxCtlMod_Cur^:=xCtlMod_Cur;
END_IF
IF i_pbyWaitCnt<>0 THEN
	i_pbyWaitCnt^:=byWaitCnt;
END_IF

(* ---- KS_ReDealCtlCommand.st ---- *)
(*@CES
Name=KS_ReDealCtlCommand
Type=FunctionBlock
TypeGuid=6f9dac99-8de1-4efc-8465-68ac443b7d08
Guid=29a1e171-811f-44f6-94ab-28798cfe2ff0
HasDeclaration=True
HasImplementation=True
*)
{DECLARATION}
FUNCTION KS_ReDealCtlCommand : BOOL
(*重新处理控制命令@因为位置模式有最大值的限制,这里将位置模式的控制拆分为先速度模式在位置模式输出控制*)
VAR_INPUT
	i_pstStInkGrooveCtl:POINTER TO StInkGrooveCtl;(*输入的控制命令*)
	i_byPulseOutSts: BYTE;(*反馈的输出状态|=0 不输出|=1 输出@逻辑|=2反馈正在运行|=3异常|=255 准备写入@进入case*)
	i_pbyPosModeSts:POINTER TO BYTE;(*位置模式的状态机
											|=1 位置模式
											|=2 速度模式+位置模式下的速度模式
											|=3 取消输出使能
											|=10切换为位置模式
											|=100等待结束
									*)

	i_pxPulseOutEn:POINTER TO BOOL;(*使能输出*)
	i_pxMoveDir:POINTER TO BOOL;(*运动方向*)
	i_pxPulseCtlMode:POINTER TO BOOL;(*控制模式|=false速度模式|=true 位置模式*)
	i_pxVelMod_Run:POINTER TO BOOL;(*速度控制模式下|速度使能标志*)
	i_prVelMod_Vel:POINTER TO REAL;(*速度控制模式下的速度*)
	i_pwPosMod_Pulse:POINTER TO WORD;(*位置控制模式下的脉冲数*)
	i_pxPosMod_InPos:POINTER TO BOOL;(*位置模式到位标志*)
END_VAR
VAR
	pstStInkGrooveCtl: POINTER TO StInkGrooveCtl;
	byPosModeSts: BYTE;(*位置模式的状态机	|=1 位置模式
											|=2 速度模式+位置模式下的速度模式
											|=3 取消输出使能
											|=10切换为位置模式
											|=100等待结束
								*)
	(*脉冲控制函数需要的输入处理@用于处理1色*)
	xPulseOutEn:BOOL;(*脉冲输出使能*)
	iPulseOutState:TypeEnumStepDriveStat;(*脉冲控制状态@状态机标志*)
(*	wLastPulse_Act_Rd_PulseOut: WORD;(*备份实际脉冲值*)*)
	byOutSts: BYTE;(*反馈的输出状态|=0 不输出|=1 输出@逻辑|=2反馈正在运行|=3异常|=255 准备写入@进入case*)
(*	xCtlMod_Cur: BOOL;(*当前的控制模式*)*)
	xVelMod_Run: BOOL;(*速度模式.控制使能标志*)
	xCtlMode: BOOL;(*控制模式*)
	rSetVel: REAL;(*速度模式的速度*)
	wSetPulse:WORD;(*设置的脉冲*)
	xMoveDir: BOOL;(*运动的方向*)
	diDeltaPulse: DINT;
	xInPos: BOOL;(*位置到位*)
(*	wNeedMovePulse: WORD;(*需要运动的脉冲@不清除*)*)
END_VAR
{IMPLEMENTATION}
IF i_pbyPosModeSts<>0 THEN
	byPosModeSts:=i_pbyPosModeSts^;
END_IF
IF i_pwPosMod_Pulse<>0 THEN
	wSetPulse:=i_pwPosMod_Pulse^;
END_IF
(*对于速度模式和位置模式做一些处理*)
(*对使能和控制方式做了重新处理*)
pstStInkGrooveCtl:= i_pstStInkGrooveCtl;
byOutSts:=i_byPulseOutSts;
IF pstStInkGrooveCtl^.byMovingSts<>0  THEN(*可以运动了*)
	xMoveDir:=pstStInkGrooveCtl^.xMoveDir;
	rSetVel:=pstStInkGrooveCtl^.rVel;
	xVelMod_Run:=FALSE;
	IF pstStInkGrooveCtl^.xCtlMode THEN(*位置模式的时候|按照速度模式+位置模式实现*)
		CASE byPosModeSts OF
			0:
				(*判断留点余量*)
				IF ABS(pstStInkGrooveCtl^.diMoveDis_Pulse)<65000(*65535*) THEN(*未超限|直接使用位置模式模块位置模式最大65535脉冲*)
					byPosModeSts:=1;
				ELSE
					byPosModeSts:=2;
				END_IF
				wSetPulse:=0;(*设置的脉冲值先写0*)
			1:(*位置模式*)
				xPulseOutEn:=TRUE;
				xCtlMode:=TRUE;(*按照位置模式*)
				wSetPulse:=DINT_TO_WORD(pstStInkGrooveCtl^.diMoveDis_Pulse);
(*				wNeedMovePulse:=wSetPulse;*)
				byPosModeSts:=100;
			2:(*速度模式+位置模式下的速度模式*)
				xPulseOutEn:=TRUE;
				xCtlMode:=FALSE;
				xVelMod_Run:=TRUE;
				diDeltaPulse:=ABS(pstStInkGrooveCtl^.diMoveDis_Pulse)-ABS(pstStInkGrooveCtl^.diThisMovedPulse);
				IF (diDeltaPulse<65535 AND diDeltaPulse>0) THEN
					byPosModeSts:=3;(*先退出速度模式再进入位置模式*)
				ELSIF diDeltaPulse<0 THEN
					byPosModeSts:=110;(*直接结束吧*)
					xInPos:=TRUE;(*到位标志*)
				ELSE
					IF byOutSts=3 THEN(*速度模式运动异常*)
						byPosModeSts:=110;(*直接结束吧*)
						xInPos:=TRUE;(*到位标志*)
					END_IF
				END_IF
			3:(*退出速度模式*)
				xPulseOutEn:=FALSE;
				IF byOutSts=0 OR byOutSts=3 THEN(*停止运动了*)
					IF byOutSts=0 THEN
						byPosModeSts:=10;(*重新进入位置模式*)
					ELSE(*速度模式运动长时间没反应*)
						byPosModeSts:=110;
						xInPos:=TRUE;(*到位标志*)
					END_IF
				END_IF
			10:(*后半程进入位置模式\并未退出运动控制case@本次运动脉冲不会清除*)
				xPulseOutEn:=TRUE;
				xCtlMode:=TRUE;(*按照位置模式*)
				diDeltaPulse:=ABS(pstStInkGrooveCtl^.diMoveDis_Pulse)-ABS(pstStInkGrooveCtl^.diThisMovedPulse);
				IF diDeltaPulse>65535 THEN
					diDeltaPulse:=65535;
				ELSIF diDeltaPulse>0 THEN;
				ELSE
					diDeltaPulse:=0;
				END_IF
				wSetPulse:=DINT_TO_WORD(diDeltaPulse);
				byPosModeSts:=100;

			100:(*等待结束*)
				xPulseOutEn:=TRUE;
				xCtlMode:=TRUE;(*按照位置模式*)
				IF ABS(pstStInkGrooveCtl^.diThisMovedPulse) >= ABS(pstStInkGrooveCtl^.diMoveDis_Pulse) THEN(*本次运动的超过了需要运动的*)
					byPosModeSts:=110;
					xInPos:=TRUE;(*到位标志*)
				END_IF
			110:(*到位了*)
				xInPos:=TRUE;(*到位标志*)
		ELSE
			byPosModeSts:=0;
(*			wNeedMovePulse:=0;*)
			wSetPulse:=0;
		END_CASE
	ELSE(*速度模式*)
		wSetPulse:=0;(*设置的脉冲值先写0*)
		byPosModeSts:=0;
		xPulseOutEn:=TRUE;
		xCtlMode:=FALSE;
		(*速度模式,停止就减速停吧*)
		xVelMod_Run:=TRUE;
	END_IF
ELSE(*停止运动了*)
	byPosModeSts:=0;
	wSetPulse:=0;(*设置的脉冲值先写0*)
END_IF

IF i_pbyPosModeSts<>0 THEN
	i_pbyPosModeSts^:=byPosModeSts;
END_IF
IF i_pxPulseOutEn<>0 THEN
	i_pxPulseOutEn^:=xPulseOutEn;
END_IF
IF i_pxMoveDir<>0 THEN
	i_pxMoveDir^:=xMoveDir;
END_IF
IF i_pxPulseCtlMode<>0 THEN
	i_pxPulseCtlMode^:=xCtlMode;
END_IF
IF i_pxVelMod_Run<>0 THEN
	i_pxVelMod_Run^:=xVelMod_Run;
END_IF
IF i_prVelMod_Vel<>0 THEN
	i_prVelMod_Vel^:=rSetVel;
END_IF
IF i_pwPosMod_Pulse<>0 THEN
	i_pwPosMod_Pulse^:=wSetPulse;
END_IF
IF i_pxPosMod_InPos<>0 THEN
	i_pxPosMod_InPos^:=xInPos;
END_IF

(* ---- KS_FB_InkGrooveCtl.st ---- *)
(*@CES
Name=KS_FB_InkGrooveCtl
Type=FunctionBlock
TypeGuid=6f9dac99-8de1-4efc-8465-68ac443b7d08
Guid=49f5b0cb-8423-4005-950e-682392de8c5e
HasDeclaration=True
HasImplementation=True
*)
{DECLARATION}
FUNCTION_BLOCK KS_FB_InkGrooveCtl
(*油墨槽升降功能块@控制1色(使用模块控制输出)*)
(*1色为主站时使用该功能块控制模块输出@目前还没支持io输出*)
VAR_INPUT
	i_xEn							: BOOL;(*功能块使能*)
	i_xCanMove						: BOOL;(*可以运动标志@例如非急停*)
	(*脉冲控制参数@主要用于1色为主站时的控制*)
	i_xMoveDirRev					: BOOL;(*方向取反*)
	i_dwPulse_1r					: DWORD;(*一圈的脉冲数*)
	i_rDis_1Pulse 					: REAL; (*单位脉冲距离mm/p*)
	i_iVel_Sa						: INT;(*脉冲输出的启动速度|r/min*)
	i_iSetVel 						: INT;(*运动速度|r/min*)
	i_iAccTime_ms					: INT;(*脉冲加速时间@100*)(*ms*)
	i_iMaxMoveDis					: INT;(*最大运动距离@mm*)
(*
	(*反馈参数@模块方式控制*)
	i_wPulse_Act_Rd_1U 				: WORD ; (*1色控制的脉冲输出值*)
	i_xPulseOutting_Rd_1U			: BOOL; (*1色控制的运动中标志*)
*)
	(*轴信息*)
	i_iGrpAxisNum_Pu						: INT; (*色组轴数*)
	i_aiGrpAxisList							: ARRAY [1..MAX_STATION_NUM] OF INT; (*系的轴列表*)
	i_auiStationTypeID						: ARRAY [0..MAX_STATION_NUM] OF UINT;(*驱动器类型字|索引为站号*)
	i_pastStAxisParam						: POINTER TO ARRAY [1..MAX_STATION_NUM] OF StAxisParam;
	i_pastStIOMap_AxisBasic					: POINTER TO ARRAY [1..MAX_STATION_NUM] OF StIOMap_AxisBasic;
	i_pstInkGrooveInf_1U_Module				: POINTER TO StDigitalMicroStepDrive;(*模块方式下获取信息和写入信息*)
END_VAR
VAR_OUTPUT
	o_xEn:BOOL;
	o_xUseControllerIO_1U: BOOL;(*1色使用控制器io@逻辑还未实现1色按照驱动器io输出|1色控制默认使用模块输出*)
	o_stStPulseModuleInf_Wr_1U: StPulseModuleInf_Wr;(*主要是1色按照模块方式输出*)
END_VAR
VAR
	in: INT;
	iAxisId:INT;
	xClrMsg: BOOL;(*提示信息清除*)
	pstStAxisParam:POINTER TO StAxisParam;
	pstStIOMap_AxisBasic:POINTER TO StIOMap_AxisBasic;
	(*共享内存里的数据@测试还未替换*)
	(*功能块中的变量*)
	pstStInkGrooveCtl:POINTER TO StInkGrooveCtl;(*油墨槽控制参数结构体*)
	xInPos: BOOL;(*位置到位*)

	(*1色使用模块方式控制的变量*)
	xPulseOutEn_1U:BOOL;(*脉冲输出使能*)
	xInPos_1U: BOOL;(*位置到位@本地控制的*)
	xVelMod_Run_1U: BOOL;(*速度模式.控制使能标志*)
	xCtlMode_1U: BOOL;(*控制模式*)
	rSetVel_1U: REAL;(*速度模式的速度*)
	xMoveDir_1U: BOOL;(*运动的方向*)
	byPosModeSts_1U: BYTE;(*位置模式的状态机	|=1 位置模式
											|=2 速度模式+位置模式下的速度模式
											|=3 取消输出使能
											|=10切换为位置模式
											|=100等待结束
								*)
	byPulseOutSts_1U: BYTE;(*输出状态|=0 不输出|=1 输出@逻辑|=2反馈正在运行|=3异常|=255 准备写入@进入case*)
	wNeedMovePulse_1U: WORD;(*需要运动的脉冲@不清除*)
	wPrevNeedMovePulse_1U: WORD;
	wSetPulse_1U:WORD;(*设置的脉冲数@获取后会清除*)
	(*模块脉冲控制输出*)
	xCtlMod_Cur_1U: BOOL;(*当前的控制模式*)
	iPulseOutState_1U:TypeEnumStepDriveStat;(*脉冲控制状态@状态机标志*)
	diThisMovePulse_1U: DINT;(*本地控制本次运动的脉冲@1色*)
	wLastPulse_Act_Rd_PulseOut: WORD;(*备份实际脉冲值*)
	byWaitCnt: BYTE;(*计时计数值*)
	(*反馈参数@模块方式控制*)
	wPulse_Act_Rd_1U 				: WORD ; (*1色控制的脉冲输出值*)
	xPulseOutting_Rd_1U			: BOOL; (*1色控制的运动中标志*)

	(*上升*)
	xClick_InkGroove_Up : BOOL ;	(*上升单击事件*)
	xDoubleClick_InkGroove_Up : BOOL ;(*上升双击事件*)
	xHold_InkGroove_Up : BOOL ;(*上升长按事件*)
	awCnt_InkGroove_Up : ARRAY [1..16] OF WORD ;(*上升状态*)

	(*下降*)
	xClick_InkGroove_Dn : BOOL ;	(*下降单击事件*)
	xDoubleClick_InkGroove_Dn : BOOL ;(*下降双击事件*)
	xHold_InkGroove_Dn : BOOL ;(*下降长按事件*)
	awCnt_InkGroove_Dn : ARRAY [1..16] OF WORD ;(*下降状态*)
	wPulse_Act_Rd: WORD;
	xMoving_Act: BOOL;(*实际运动中标志*)
	iStationId: INT;(*站号*)
	xCtlEn: BOOL;(*2025.6.6.114812 控制使能标志*)
	xIsMaster_1U: BOOL;(*1色是主站*)
	xUseModule: BOOL;(*使用过模块标志@用来清理数据*)
	xVelMode_MoveFailed: BOOL;(*速度模式运动失败*)
END_VAR
{IMPLEMENTATION}
IF i_pstInkGrooveInf_1U_Module<>0 AND
	i_pastStIOMap_AxisBasic<>0 AND
	i_pastStAxisParam<>0 THEN;
ELSE
	RETURN;
END_IF
(*动作控制@所有轴(1--16)*)
(*模块控制的时候获取反馈数据*)
IF o_xUseControllerIO_1U AND FALSE THEN(*还未实现|先强制false*)
	;
ELSE
	wPulse_Act_Rd_1U:=i_pstInkGrooveInf_1U_Module^.wStepDrivePulse_Act_Rd;
	xPulseOutting_Rd_1U:=i_pstInkGrooveInf_1U_Module^.xStepDriveWorking;
END_IF

xIsMaster_1U:=FALSE;
FOR in:=1 TO i_iGrpAxisNum_Pu BY 1 DO
	iAxisId:=i_aiGrpAxisList[in];
	IF iAxisId>0 AND iAxisId<=16 THEN
		pstStAxisParam:=ADR(i_pastStAxisParam^[iAxisId]);
		pstStIOMap_AxisBasic:=ADR(i_pastStIOMap_AxisBasic^[iAxisId]);
		pstStInkGrooveCtl:= ADR(pstStAxisParam^.stStInkGrooveCtl);
		iStationId:=pstStAxisParam^.iStationId;

		(*检查驱动器是不是支持|确认使能标志*)
		xCtlEn:=i_xEn;(*初始化为使能输入*)
		IF iStationId>=0 AND iStationId<=MAX_STATION_NUM THEN
			IF iStationId<>0 THEN(*从站*)
				IF i_auiStationTypeID[iStationId] = CONTROLLER_GTSD16D_AIO OR(*新款16d-1*)
					i_auiStationTypeID[iStationId] = CONTROLLER_GTSD16D_AIO_ISO OR(*新款16d-2*)
					i_auiStationTypeID[iStationId] = CONTROLLER_GTSD16M_AIO THEN(*新款16m*)

					IF iAxisId=1 THEN(*1#轴@从站*)
						o_xUseControllerIO_1U:=TRUE;
					END_IF
				ELSE
					xCtlEn:=FALSE;
					IF iAxisId=1 THEN(*1#轴@从站*)
						o_xUseControllerIO_1U:=FALSE;
					END_IF
				END_IF
			ELSE(*主站@肯定是色组轴|else里的逻辑可有可无*)
				IF iAxisId=1 THEN(*1#轴*)
					xIsMaster_1U:=TRUE;
					IF i_auiStationTypeID[iStationId] = CONTROLLER_GTSD16M_AIO THEN(*新款16m*)
						o_xUseControllerIO_1U:=TRUE;
					ELSE
						o_xUseControllerIO_1U:=FALSE;
					END_IF
				ELSE(*非1#轴就不理*)
					xCtlEn:=FALSE;
					o_xUseControllerIO_1U:=FALSE;
				END_IF
			END_IF
		END_IF

		(*一些反馈标志处理,有本地信息也有通讯讯息*)
		IF xCtlEn THEN(*使能了*)
			(*将保持的值写入到油墨槽变量|下面逻辑会继续更新*)
			pstStInkGrooveCtl^.diPulse_Moved:=pstStAxisParam^.diPulseValue_16D;
			IF iAxisId=1 THEN
				IF xIsMaster_1U THEN(*1色是主站@反馈信息都从本地获取*)
					xMoving_Act:=byPulseOutSts_1U<>0;
					wPulse_Act_Rd:=wPulse_Act_Rd_1U;
					xVelMode_MoveFailed:=byPulseOutSts_1U=3;
					xInPos:=xInPos_1U;
				ELSE(*不是主站|通讯获取*)
					xMoving_Act:=pstStAxisParam^.xPulse_Outing_16D;(*因为是通讯获取的，能不能可靠拿到标志|要注意*)
					wPulse_Act_Rd:=pstStAxisParam^.wPulse_Rd_16D;
					xVelMode_MoveFailed:=pstStAxisParam^.byInkGroovePulseOutSts = 3;
					xInPos:=pstStAxisParam^.xInkGroove_InPos;
				END_IF
			ELSE(*其他色组通讯获取信息|*)
				xMoving_Act:=pstStAxisParam^.xPulse_Outing_16D;
				wPulse_Act_Rd:=pstStAxisParam^.wPulse_Rd_16D;
				xVelMode_MoveFailed:=pstStAxisParam^.byInkGroovePulseOutSts = 3;
				xInPos:=pstStAxisParam^.xInkGroove_InPos;
			END_IF
		ELSE(*不使能*)
			xMoving_Act:=FALSE;
			wPulse_Act_Rd:=0;
			xVelMode_MoveFailed:=FALSE;
			xInPos:=TRUE;
		END_IF

		(*io处理*)
		IF NOT xCtlEn OR NOT i_xCanMove THEN
			pstStIOMap_AxisBasic^.i_xBtnInkGroove_Up:=FALSE;
			pstStIOMap_AxisBasic^.i_xBtnInkGroove_Dn:=FALSE;
		END_IF

		KS_BtnClick(
			pstStIOMap_AxisBasic^.i_xBtnInkGroove_Up(*i_xBtn*),(*上升信号*)
			300(*i_wTime_ms*),
			INT_TO_BYTE(gc_iCycleTime_Plc)(*i_byCycleTime_ms*),
			ADR(xClick_InkGroove_Up)(*i_pxClick*),
			ADR(xDoubleClick_InkGroove_Up)(*i_pxDoubleClick*),
			ADR(xHold_InkGroove_Up)(*i_pxHold*),
			ADR(awCnt_InkGroove_Up[iAxisId])(*i_pwCnt*));

		KS_BtnClick(
			pstStIOMap_AxisBasic^.i_xBtnInkGroove_Dn(*i_xBtn*),(*上升信号*)
			300(*i_wTime_ms*),
			INT_TO_BYTE(gc_iCycleTime_Plc)(*i_byCycleTime_ms*),
			ADR(xClick_InkGroove_Dn)(*i_pxClick*),
			ADR(xDoubleClick_InkGroove_Dn)(*i_pxDoubleClick*),
			ADR(xHold_InkGroove_Dn)(*i_pxHold*),
			ADR(awCnt_InkGroove_Dn[iAxisId])(*i_pwCnt*));

		KS_InkGrooveCtl_1Axis(
			xCtlEn(*i_xEn*),
			i_xCanMove(*i_xCanMove*),
			xClrMsg(*i_xClrMsg*),
			i_rDis_1Pulse(*i_lrDis_1Pulse*),
			INT_TO_BYTE(gc_iCycleTime_Plc)(*i_iCycleTime_Plc*),
			pstStAxisParam^.lrGirth(*i_rGirth*),
			pstStAxisParam^.xInkGroove_BaseInfValid(*i_xBaseInfValid*),
			pstStAxisParam^.rInkGroove_Girth_Base(*i_rGirth_Base*),
			pstStAxisParam^.rInkGroove_Pos_Base(*i_rPos_Base*),
			i_xMoveDirRev(*i_xMoveDirRev*),
			xHold_InkGroove_Up(*i_xUp*),
			pstStIOMap_AxisBasic^.i_xInkGrooveUplimt(*i_xUplimt*),
			xHold_InkGroove_Dn(*i_xDn*),
			xDoubleClick_InkGroove_Dn(*i_xDn_Auto*),
			pstStIOMap_AxisBasic^.i_xInkGrooveDnlimt(*i_xDnlimt*),
			xClick_InkGroove_Up, (*i_xUpClick*)
			xClick_InkGroove_Dn,(*i_xDnClick *)
			xDoubleClick_InkGroove_Up (*i_xToTarPos_Auto*),
			pstStIOMap_AxisBasic^.i_xInkGrooveDnlimt(*i_xZeroSig*),
			INT_TO_REAL(i_iSetVel)(*i_rSetVel*),
			INT_TO_REAL(i_iMaxMoveDis)(*i_rMaxMoveDis*),
			wPulse_Act_Rd(*i_wPulse_Act_Rd*),(*反馈*)
			xInPos(*i_xInPos*),(*反馈*)
			xMoving_Act(*i_xMoving_Act*),(*反馈*)
			xVelMode_MoveFailed(*i_xVelMode_MoveFailed*),
			pstStInkGrooveCtl(*i_pstStInkGrooveCtl*));

		(*获取自动的基础信息@1-16色*)
		KS_GetInkGrooveBaseInf(
			pstStInkGrooveCtl^.xZeroValid(*i_xEn*),
			pstStAxisParam^.xGetInkGoove_BaseInf(*i_xGetBtn*),
			pstStAxisParam^.lrGirth(*i_rGirth*),
			pstStInkGrooveCtl^.rPos_Cur(*i_rPos_Cur*),
			ADR(pstStAxisParam^.xInkGroove_BaseInfValid)(*i_pxBaseInfValid*),
			ADR(pstStAxisParam^.rInkGroove_Girth_Base)(*i_prGirth_Base*),
			ADR(pstStAxisParam^.rInkGroove_Pos_Base)(*i_prPos_Base*));
		pstStAxisParam^.xGetInkGoove_BaseInf:=FALSE;(*按钮复位*)

		(*从站通讯内容写入@2025.6.11.192921*)
		IF xCtlEn THEN(*使能了|处理通讯写入*)
			IF pstStInkGrooveCtl^.xCtlMode THEN(*位置模式*)
				pstStAxisParam^.wPulseCtlInf_16D:=REAL_TO_WORD(ABS(pstStInkGrooveCtl^.rMoveDis*100));
			ELSE(*速度模式*)
				pstStAxisParam^.wPulseCtlInf_16D:=REAL_TO_WORD(ABS(pstStInkGrooveCtl^.rVel*10));
			END_IF
			pstStAxisParam^.wPulse_1r_16D:=DWORD_TO_WORD(i_dwPulse_1r);
			pstStAxisParam^.byPulseCtl_DisPerPulse_16D:=REAL_TO_BYTE(i_rDis_1Pulse*100000);(*单位0.01um*)
			pstStAxisParam^.byPulseCtlBit_16D:=0;
			pstStAxisParam^.byPulseCtlBit_16D.0:=xCtlEn;(*使能@从站io才可以按照脉冲输出*)
			pstStAxisParam^.byPulseCtlBit_16D.1:=pstStInkGrooveCtl^.bySts<>0;(*运动使能*)
			pstStAxisParam^.byPulseCtlBit_16D.2:=pstStInkGrooveCtl^.xMoveDir;(*运动方向*)
			pstStAxisParam^.byPulseCtlBit_16D.3:=pstStInkGrooveCtl^.xCtlMode;(*控制模式*)
			pstStAxisParam^.diPulseValue_16D:=pstStInkGrooveCtl^.diPulse_Moved;(*已经运动的距离写入到保持变量里*)
		ELSE(*不使能*)
			IF pstStAxisParam^.byPulseCtlBit_16D.0 THEN(*作为取消使能清零的条件|在使能时候该bit会被置位*)
				pstStAxisParam^.byPulseCtlBit_16D:=0;
				pstStAxisParam^.wPulseCtlInf_16D:=0;
				pstStAxisParam^.diPulseValue_16D:=0;
			END_IF
		END_IF

	ELSE(*控制不使能*)
		;
	END_IF
END_FOR

(*模块写入信息处理@1色*)
(*对于速度模式和位置模式做一些处理*)
(*对使能和控制方式做了重新处理*)
pstStAxisParam:=ADR(i_pastStAxisParam^[1]);
pstStInkGrooveCtl:= ADR(pstStAxisParam^.stStInkGrooveCtl);
KS_ReDealCtlCommand(
	pstStInkGrooveCtl(*i_pstStInkGrooveCtl*),
	byPulseOutSts_1U(*i_byPulseOutSts*),
	ADR(byPosModeSts_1U)(*i_pbyPosModeSts*),
	ADR(xPulseOutEn_1U)(*i_pxPulseOutEn*),
	ADR(xMoveDir_1U)(*i_pxMoveDir*),
	ADR(xCtlMode_1U)(*i_pxPulseCtlMode*),
	ADR(xVelMod_Run_1U)(*i_pxVelMod_Run*),
	ADR(rSetVel_1U)(*i_prVelMod_Vel*),
	ADR(wNeedMovePulse_1U)(*i_pwPosMod_Pulse*),
	ADR(xInPos_1U)(*i_pxPosMod_InPos*));
(*设置的脉冲数@变为非0,写入到控制模块脉冲输出的函数变量*)
IF wSetPulse_1U=0 AND
	wNeedMovePulse_1U<>0 THEN
	wSetPulse_1U:=wNeedMovePulse_1U;(*wSetPulse_1U 由KS_PulseOutCtl清零*)
END_IF

IF o_xUseControllerIO_1U AND FALSE THEN(*1色使用驱动器io@还未实现-强制无效*)

	IF xUseModule THEN
		xUseModule:=FALSE;
		SysMemSet(ADR(o_stStPulseModuleInf_Wr_1U),0,SIZEOF(o_stStPulseModuleInf_Wr_1U));
		SysMemSet(ADR(i_pstInkGrooveInf_1U_Module^),0,SIZEOF(i_pstInkGrooveInf_1U_Module^));
		wLastPulse_Act_Rd_PulseOut:=wPulse_Act_Rd_1U;
		iPulseOutState_1U:=STEPDRIVE_IDLE;
		wSetPulse_1U:=0;
		diThisMovePulse_1U:=0;
		byPulseOutSts_1U:=0;
		byWaitCnt:=0;
	END_IF
ELSE(*1色使用模块*)
	(*模块控制脉冲*)
	KS_PulseOutCtl(
		xPulseOutEn_1U(*i_xEn*),
		FALSE(*i_xClrPulse_Act_Rd*),
		10(*i_byJudgeOutsts_WaitNum*),
		i_dwPulse_1r(*i_dwPulse_1r*),
		xCtlMode_1U(*i_xCtlMode*),
		xVelMod_Run_1U(*i_xVelMod_Run*),
		xMoveDir_1U(*i_xDir*),
		INT_TO_REAL(i_iVel_Sa)(*i_rVel_Sa*),
		rSetVel_1U(*i_rVel*),
		i_iAccTime_ms(*i_iAccTime_ms*),
		ADR(wSetPulse_1U)(*i_pwPulse*),
		xPulseOutting_Rd_1U(*i_xPulseOutting_Rd*),
		wPulse_Act_Rd_1U(*i_wPulse_Act_Rd*),
		ADR(iPulseOutState_1U)(*i_piState*),
		ADR(o_stStPulseModuleInf_Wr_1U.wCTL)(*i_pwCtlBit_Wr*),
		ADR(o_stStPulseModuleInf_Wr_1U.wPulseFre_Sa_Wr)(*i_pwFre_Sa_Wr*),
		ADR(o_stStPulseModuleInf_Wr_1U.wPulseFre_Tar_Wr)(*i_pwFreq_Tar_Wr*),
		ADR(o_stStPulseModuleInf_Wr_1U.wAcc_SaToTar_Wr)(*i_pwAccSaToTar_Wr*),
		ADR(o_stStPulseModuleInf_Wr_1U.wPulse_Wr)(*i_pwPulse_Pos_Wr*),
		ADR(diThisMovePulse_1U)(*i_pdiPluse_Act*),
		ADR(wLastPulse_Act_Rd_PulseOut)(*i_pwLastPulse_Act_Rd*),
		ADR(byPulseOutSts_1U)(*i_pbyOutSts*),
		ADR(xCtlMod_Cur_1U)(*i_pxCtlMod_Cur*),
		ADR(byWaitCnt)(*i_pbyWaitCnt*));

	(*写入到原来做的模块输出的结构体中去，代码好实现一些*)
	i_pstInkGrooveInf_1U_Module^.wStepDriveCTL:=o_stStPulseModuleInf_Wr_1U.wCTL;
	i_pstInkGrooveInf_1U_Module^.wStepDrivePulseFre_Sa_Wr:=o_stStPulseModuleInf_Wr_1U.wPulseFre_Sa_Wr;
	i_pstInkGrooveInf_1U_Module^.wStepDrivePulseFre_Tar_Wr:=o_stStPulseModuleInf_Wr_1U.wPulseFre_Tar_Wr;
	i_pstInkGrooveInf_1U_Module^.wStepDriveAcc_SaToTar_Wr:=o_stStPulseModuleInf_Wr_1U.wAcc_SaToTar_Wr;
	i_pstInkGrooveInf_1U_Module^.wStepDrivePulse_Wr:=o_stStPulseModuleInf_Wr_1U.wPulse_Wr;
	xUseModule:=TRUE;
END_IF
